// Mitsubishi GX Works2 project: 공개3번(FX)   PLC: FX3U/FX3UC

PROGRAM MAIN
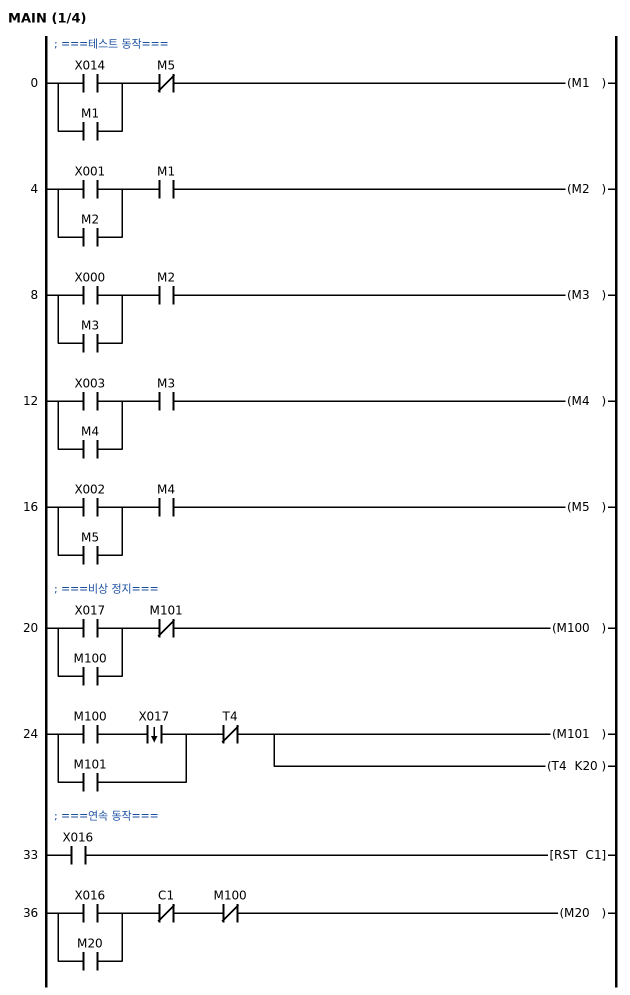
; ===테스트 동작===
0     LD      X014
      OR      M1
      ANI     M5
      OUT     M1
4     LD      X001
      OR      M2
      AND     M1
      OUT     M2
8     LD      X000
      OR      M3
      AND     M2
      OUT     M3
12    LD      X003
      OR      M4
      AND     M3
      OUT     M4
16    LD      X002
      OR      M5
      AND     M4
      OUT     M5
; ===비상 정지===
20    LD      X017
      OR      M100
      ANI     M101
      OUT     M100
24    LD      M100
      ANDF    X017
      OR      M101
      ANI     T4
      OUT     M101
      OUT     T4 K20
; ===연속 동작===
33    LD      X016
      RST     C1
36    LD      X016
      OR      M20
      ANI     C1
      ANI     M100
      OUT     M20
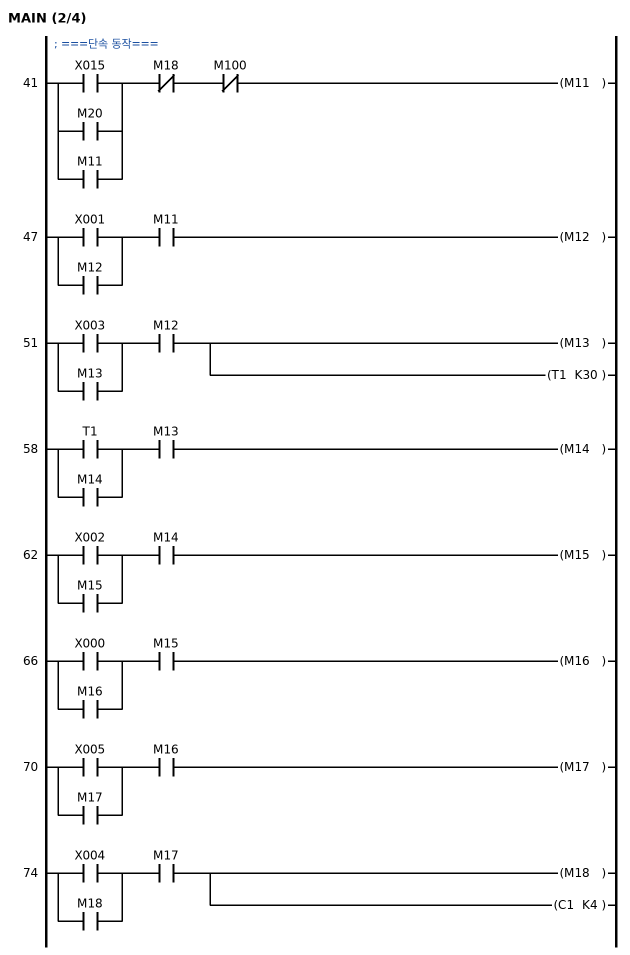
; ===단속 동작===
41    LD      X015
      OR      M20
      OR      M11
      ANI     M18
      ANI     M100
      OUT     M11
47    LD      X001
      OR      M12
      AND     M11
      OUT     M12
51    LD      X003
      OR      M13
      AND     M12
      OUT     M13
      OUT     T1 K30
58    LD      T1
      OR      M14
      AND     M13
      OUT     M14
62    LD      X002
      OR      M15
      AND     M14
      OUT     M15
66    LD      X000
      OR      M16
      AND     M15
      OUT     M16
70    LD      X005
      OR      M17
      AND     M16
      OUT     M17
74    LD      X004
      OR      M18
      AND     M17
      OUT     M18
      OUT     C1 K4
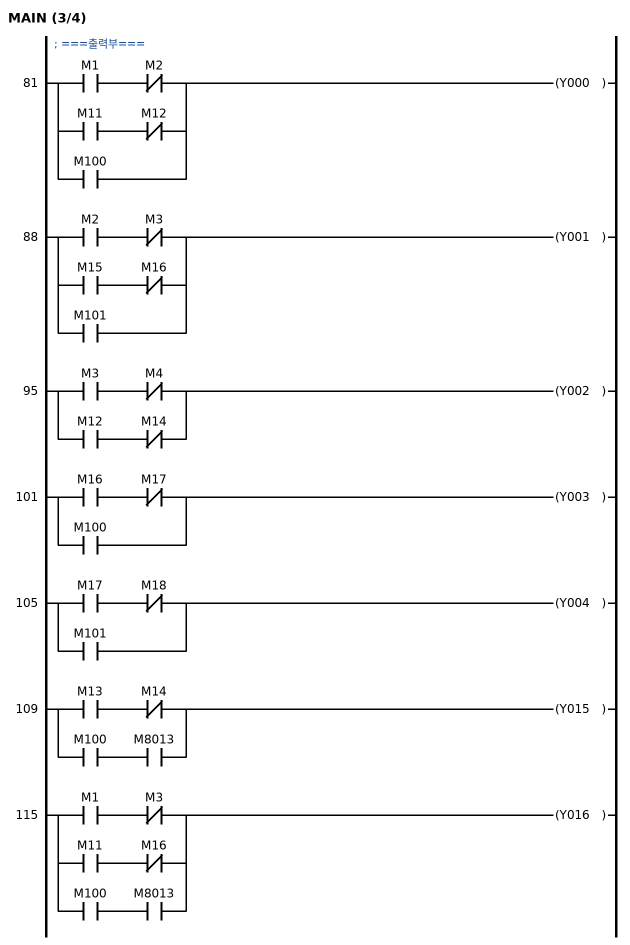
; ===출력부===
81    LD      M1
      ANI     M2
      LD      M11
      ANI     M12
      ORB
      OR      M100
      OUT     Y000
88    LD      M2
      ANI     M3
      LD      M15
      ANI     M16
      ORB
      OR      M101
      OUT     Y001
95    LD      M3
      ANI     M4
      LD      M12
      ANI     M14
      ORB
      OUT     Y002
101   LD      M16
      ANI     M17
      OR      M100
      OUT     Y003
105   LD      M17
      ANI     M18
      OR      M101
      OUT     Y004
109   LD      M13
      ANI     M14
      LD      M100
      AND     M8013
      ORB
      OUT     Y015
115   LD      M1
      ANI     M3
      LD      M11
      ANI     M16
      ORB
      LD      M100
      AND     M8013
      ORB
      OUT     Y016
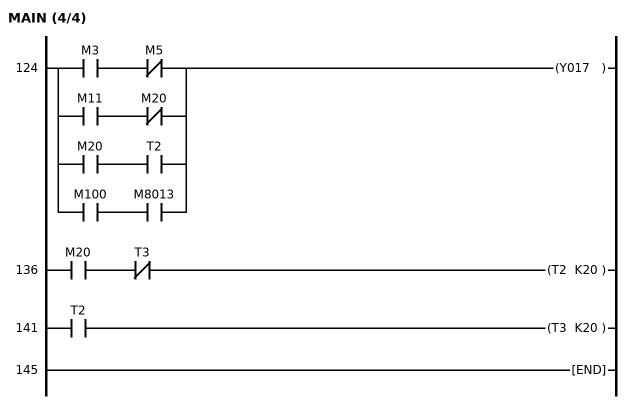
124   LD      M3
      ANI     M5
      LD      M11
      ANI     M20
      ORB
      LD      M20
      AND     T2
      ORB
      LD      M100
      AND     M8013
      ORB
      OUT     Y017
136   LD      M20
      ANI     T3
      OUT     T2 K20
141   LD      T2
      OUT     T3 K20
145   END
END_PROGRAM
